(* IEC 61131-3 sources: iolistgen/tests_support/pl_stub/src/DUTs/Valve, 7 files *)

(* ---- E_ValveAlarm.dut.st ---- *)
// Назначение: заглушка plc-process-lib 1.0.0 для проверки типов сгенерированного кода без CODESYS
//             (API.md, раздел 4.1); не библиотека — тел и внутренних переменных нет
// Автор:      kr0nsch
// Версия:     1.0.0 (выпуск библиотеки)
// Документ:   docs/GENERATORS.md, раздел «Проверка ST без CODESYS»
{attribute 'qualified_only'}
TYPE E_ValveAlarm :
(
    FailToOpen := 0,
    FailToClose := 1,
    BothLimits := 2,
    PositionLost := 3,
    TorqueTrip := 4,
    ExtFault := 5,
    InterlockAct := 6
) UINT;
END_TYPE

(* ---- E_ValveSafePos.dut.st ---- *)
// Назначение: заглушка plc-process-lib 1.0.0 для проверки типов сгенерированного кода без CODESYS
//             (API.md, раздел 15.1); не библиотека — тел и внутренних переменных нет
// Автор:      kr0nsch
// Версия:     1.0.0 (выпуск библиотеки)
// Документ:   docs/GENERATORS.md, раздел «Проверка ST без CODESYS»
{attribute 'qualified_only'}
{attribute 'strict'}
TYPE E_ValveSafePos :
(
    Closed := 0,
    Open := 1,
    Stay := 2
) INT;
END_TYPE

(* ---- E_ValveState.dut.st ---- *)
// Назначение: заглушка plc-process-lib 1.0.0 для проверки типов сгенерированного кода без CODESYS
//             (API.md, раздел 15.1); не библиотека — тел и внутренних переменных нет
// Автор:      kr0nsch
// Версия:     1.0.0 (выпуск библиотеки)
// Документ:   docs/GENERATORS.md, раздел «Проверка ST без CODESYS»
{attribute 'qualified_only'}
{attribute 'strict'}
TYPE E_ValveState :
(
    Unknown := 0,
    Closed := 1,
    Opening := 2,
    Open := 3,
    Closing := 4,
    Intermediate := 5,
    Reversing := 6,
    Fault := 7
) INT;
END_TYPE

(* ---- E_ValveType.dut.st ---- *)
// Назначение: заглушка plc-process-lib 1.0.0 для проверки типов сгенерированного кода без CODESYS
//             (API.md, раздел 15.1); не библиотека — тел и внутренних переменных нет
// Автор:      kr0nsch
// Версия:     1.0.0 (выпуск библиотеки)
// Документ:   docs/GENERATORS.md, раздел «Проверка ST без CODESYS»
{attribute 'qualified_only'}
{attribute 'strict'}
TYPE E_ValveType :
(
    SolenoidEto := 0,
    SolenoidEtc := 1,
    Motorized := 2
) INT;
END_TYPE

(* ---- ST_ValveCfg.dut.st ---- *)
// Назначение: заглушка plc-process-lib 1.0.0 для проверки типов сгенерированного кода без CODESYS
//             (API.md, раздел 15.1); не библиотека — тел и внутренних переменных нет
// Автор:      kr0nsch
// Версия:     1.0.0 (выпуск библиотеки)
// Документ:   docs/GENERATORS.md, раздел «Проверка ST без CODESYS»
{attribute 'qualified_only'}
TYPE ST_ValveCfg :
STRUCT
    eType            : E_ValveType := E_ValveType.Motorized;
    xZsoUsed         : BOOL := TRUE;
    xZscUsed         : BOOL := TRUE;
    tTravel          : TIME := T#60S;
    tLimitFilter     : TIME := T#500MS;
    tReverse         : TIME := T#1S;
    xTorqueUsed      : BOOL := FALSE;
    xCloseOnTorque   : BOOL := FALSE;
    eSafePos         : E_ValveSafePos := E_ValveSafePos.Closed;
    wInterlockMask   : WORD := 16#FFFF;
    wPermitOpenMask  : WORD := 16#FFFF;
    wPermitCloseMask : WORD := 16#FFFF;
    tResetWindow     : TIME := T#3S;
    udiMaintCycles   : UDINT := 0;
    udiAlarmIdBase   : UDINT := 0;
    // lint:allow STL007 имя массива по контракту API.md (префикс a + тип элемента)
    astAlarm       : ARRAY[0..GVL_Const.DEV_ALARMS_MAX - 1] OF ST_AlarmCfg := [
            (ePriority := E_AlarmPriority.Medium),
            (ePriority := E_AlarmPriority.Medium),
            (ePriority := E_AlarmPriority.Medium),
            (ePriority := E_AlarmPriority.Medium),
            (ePriority := E_AlarmPriority.Medium),
            (ePriority := E_AlarmPriority.Medium),
            (ePriority := E_AlarmPriority.None),
            (ePriority := E_AlarmPriority.None)];
END_STRUCT
END_TYPE

(* ---- ST_ValveCmd.dut.st ---- *)
// Назначение: заглушка plc-process-lib 1.0.0 для проверки типов сгенерированного кода без CODESYS
//             (API.md, раздел 15.1); не библиотека — тел и внутренних переменных нет
// Автор:      kr0nsch
// Версия:     1.0.0 (выпуск библиотеки)
// Документ:   docs/GENERATORS.md, раздел «Проверка ST без CODESYS»
{attribute 'qualified_only'}
TYPE ST_ValveCmd :
STRUCT
    stCommon    : ST_DeviceCmd;
    xOpen       : BOOL;
    xClose      : BOOL;
    xStop       : BOOL;
    xResetMaint : BOOL;
END_STRUCT
END_TYPE

(* ---- ST_ValveSts.dut.st ---- *)
// Назначение: заглушка plc-process-lib 1.0.0 для проверки типов сгенерированного кода без CODESYS
//             (API.md, раздел 15.1); не библиотека — тел и внутренних переменных нет
// Автор:      kr0nsch
// Версия:     1.0.0 (выпуск библиотеки)
// Документ:   docs/GENERATORS.md, раздел «Проверка ST без CODESYS»
{attribute 'qualified_only'}
TYPE ST_ValveSts :
STRUCT
    stCommon         : ST_DeviceSts;
    eState           : E_ValveState;
    wInterlock       : WORD;
    wPermitMissing   : WORD;
    uiFirstOut       : UINT;
    uiTravelRemain_s : UINT;
    wReserve         : WORD;
    udiCycles        : UDINT;
    udiCyclesMaint   : UDINT;
    rActTime_h       : REAL;
END_STRUCT
END_TYPE
